(* IEC 61131-3 sources: SortJet_MasterSPS_Aufbau.fbsproj/09_Station/Stationen/Faecherwagen [301-305]/Basic_Faecherwagenstation_FB_V01_00_00.fb.st^, 19 files *)

(* ---- A_Changelog.act.st ---- *)
(* METADATA
{
	"v3Meta": {
		"objectGuid": "929bf022-d5bd-484d-b38d-56fc386ae04b"
	}
}
*)
{attribute 'excludefrombuild'}
ACTION A_Changelog
(* !!! VERSIONSÄNDERUNGEN WERDEN HIER DETAILLIERT DOKUMENTIERT !!!

- 2026-11-24 - V01_00_00: Tobias Brekerbohm
  - Erste Freigabe SortJet-Master
*)
END_ACTION

(* ---- A_ScheibenDeaktivierteStationMelden.act.st ---- *)
(* METADATA
{
	"v3Meta": {
		"objectGuid": "9787c6c4-89ac-4e67-aebe-436ca2600e9a"
	}
}
*)
ACTION A_ScheibenDeaktivierteStationMelden
// @TEXT_IMPLEMENTATION := 'ST'
//-------------------------------------------------------------------------------------------------
// DEAKTIVIERTE STATION: SCHEIBEN AN MMI MELDEN
//-------------------------------------------------------------------------------------------------
(* Hinweis:
   - Ersetzt die gleichnamige Aktion von Basic_Station_FB (auch beim Aufruf aus deren Rumpf)
   - Faecherwagenstationen melden dem MMI keine Scheiben auf der Station
*)
;
END_ACTION

(* ---- A_Schnittstelle.act.st ---- *)
(* METADATA
{
	"v3Meta": {
		"objectGuid": "4b006156-55f0-4052-a03b-8c052b439175"
	}
}
*)
ACTION A_Schnittstelle
//-------------------------------------------------------------------------------------------------
// SCHNITTSTELLE
//-------------------------------------------------------------------------------------------------

// Allgemeiner Teil: Auftrag aktiv, Stationsnummern, Fehler, Freigabe, Handfunktionen
SUPER^.A_Schnittstelle();

(* Hinweis:
   - Schnittstelle zwischen den Stationen [Transportkopplung]
*)
BasisStationsParameter.OutGlasTransport[cWAND_1].bEinlaufsensor         REF= bgFALSE;
BasisStationsParameter.OutGlasTransport[cWAND_1].bAuslaufsensor         REF= bgFALSE;
BasisStationsParameter.OutGlasTransport[cWAND_1].bBereitZumAustransport REF= bpOutBereitZumAustransport;
BasisStationsParameter.OutGlasTransport[cWAND_1].bBereitZumEintransport REF= bpOutBereitZumEintransport;
BasisStationsParameter.OutGlasTransport[cWAND_1].rGeschwindigkeit       REF= rgNULL;
END_ACTION

(* ---- A_Visu.act.st ---- *)
(* METADATA
{
	"v3Meta": {
		"objectGuid": "97dd6b9c-083d-47d5-ad19-d2fe11b9c8f1"
	}
}
*)
ACTION A_Visu
//-------------------------------------------------------------------------------------------------
// STATUS FUER DIE VISU
//-------------------------------------------------------------------------------------------------
// Allgemeiner Teil fuer alle Varianten; die Variante ergaenzt Faecherwagen, Lichtschranke und
// ihre Endlagen (abEndlage, Index = Bit der zugehoerigen Handfunktion)
IF PruefungWertImIntervall( BasisStationsParameter.stMKs.stStationsNummern.NummerSPS,
                            cERSTE_FAECHERWAGENSTATIONS_NR,
                            cLETZTE_FAECHERWAGENSTATIONS_NR )
THEN
  astgFaecherwagenstatusVisu[BasisStationsParameter.stMKs.stStationsNummern.NummerSPS].bBoxInHomePosition             := bpBoxInHomePosition;
  astgFaecherwagenstatusVisu[BasisStationsParameter.stMKs.stStationsNummern.NummerSPS].bStatusStationInBeladePosition := bpStatusStationInBeladePosition;
  astgFaecherwagenstatusVisu[BasisStationsParameter.stMKs.stStationsNummern.NummerSPS].bAuftragAktiv                  := bpAuftragAktiv;
  astgFaecherwagenstatusVisu[BasisStationsParameter.stMKs.stStationsNummern.NummerSPS].bFehler                        := BasisStationsParameter.bFehler;
  astgFaecherwagenstatusVisu[BasisStationsParameter.stMKs.stStationsNummern.NummerSPS].eStatus                        := eLetzterStatus;
  astgFaecherwagenstatusVisu[BasisStationsParameter.stMKs.stStationsNummern.NummerSPS].bRolltorOben                   := in_bRolltorGeoeffnet;
  astgFaecherwagenstatusVisu[BasisStationsParameter.stMKs.stStationsNummern.NummerSPS].bRolltorUnten                  := bpRolltorUnten;
  astgFaecherwagenstatusVisu[BasisStationsParameter.stMKs.stStationsNummern.NummerSPS].wRFID_Nummer                   := wlRFID_Nummer;
  astgFaecherwagenstatusVisu[BasisStationsParameter.stMKs.stStationsNummern.NummerSPS].abEndlage[5]                   := in_bRolltorGeoeffnet;
  astgFaecherwagenstatusVisu[BasisStationsParameter.stMKs.stStationsNummern.NummerSPS].abEndlage[6]                   := bpRolltorUnten;
END_IF
END_ACTION

(* ---- bAuftragAktiv.prop.st ---- *)
(* METADATA
{
	"v3Meta": {
		"objectGuid": "3a197e04-0bcd-4579-a4af-806c82b87acf",
		"subObjects": {
			"get": {
				"objectGuid": "bd81e771-6b2a-41b3-b424-5effe3645496"
			}
		}
	}
}
*)
PROPERTY_Get bAuftragAktiv : BOOL
VAR
END_VAR
bAuftragAktiv := bpAuftragAktiv;END_PROPERTY

(* ---- bBoxInHomePosition.prop.st ---- *)
(* METADATA
{
	"v3Meta": {
		"objectGuid": "9ae1053e-7eaa-4017-919c-7a919c9e2ca3",
		"subObjects": {
			"get": {
				"objectGuid": "c7a204ff-f1d2-4f02-aa57-0c1f7686d3d7"
			}
		}
	}
}
*)
PROPERTY_Get bBoxInHomePosition : BOOL
VAR
END_VAR
bBoxInHomePosition := bpBoxInHomePosition;END_PROPERTY

(* ---- bDone.prop.st ---- *)
(* METADATA
{
	"v3Meta": {
		"objectGuid": "7e3afc40-fd10-411a-82e2-c2f76dbe13b7",
		"subObjects": {
			"get": {
				"objectGuid": "a4174cb2-9640-462a-838e-1c212c18065f"
			}
		}
	}
}
*)
PROPERTY_Get bDone : BOOL
VAR
END_VAR
bDone := bpDone;END_PROPERTY

(* ---- bErzwingeAusschleusen.prop.st ---- *)
(* METADATA
{
	"v3Meta": {
		"objectGuid": "4cee021b-c5d5-4f3b-aa29-0070cbf1b16c",
		"subObjects": {
			"get": {
				"objectGuid": "1eace140-85af-4621-b197-e1bb9b84e0ab"
			}
		}
	}
}
*)
PROPERTY_Get bErzwingeAusschleusen : BOOL
VAR
END_VAR
bErzwingeAusschleusen := bpErzwingeAusschleusen;END_PROPERTY

(* ---- bErzwingeEinschleusen.prop.st ---- *)
(* METADATA
{
	"v3Meta": {
		"objectGuid": "82a9f007-64ac-4edb-aa26-a15d51300ac1",
		"subObjects": {
			"get": {
				"objectGuid": "2fa276e3-c875-4651-a2ef-8e71ffca1126"
			}
		}
	}
}
*)
PROPERTY_Get bErzwingeEinschleusen : BOOL
VAR
END_VAR
bErzwingeEinschleusen := bpErzwingeEinschleusen;END_PROPERTY

(* ---- bFehler.prop.st ---- *)
(* METADATA
{
	"v3Meta": {
		"objectGuid": "15bf96d6-b3ab-4293-98f3-daa693f44265",
		"subObjects": {
			"get": {
				"objectGuid": "7173d561-01b0-4b6a-be06-4d55a19c8095"
			}
		}
	}
}
*)
PROPERTY_Get bFehler : BOOL
VAR
END_VAR
bFehler := bpFehler;END_PROPERTY

(* ---- bMerkerEinschleusenQuittiert.prop.st ---- *)
(* METADATA
{
	"v3Meta": {
		"objectGuid": "bcf8d110-caa9-4eeb-bc74-c675be36606a",
		"subObjects": {
			"get": {
				"objectGuid": "c1b86ccc-2e67-4907-bc19-e7facae66067"
			}
		}
	}
}
*)
PROPERTY_Get bMerkerEinschleusenQuittiert : BOOL
VAR
END_VAR
bMerkerEinschleusenQuittiert := blMerkerEinschleusenQuittiert;END_PROPERTY

(* ---- bOutBereitZumAustransport.prop.st ---- *)
(* METADATA
{
	"v3Meta": {
		"objectGuid": "40e5f93b-ff00-4f78-b9f3-71c706ff1514",
		"subObjects": {
			"get": {
				"objectGuid": "2b4ba9cb-deb4-4b61-92f3-2bedee948b9f"
			}
		}
	}
}
*)
PROPERTY_Get bOutBereitZumAustransport : BOOL
VAR
END_VAR
bOutBereitZumAustransport := bpOutBereitZumAustransport;END_PROPERTY

(* ---- bOutBereitZumEintransport.prop.st ---- *)
(* METADATA
{
	"v3Meta": {
		"objectGuid": "529f8d13-9d58-45ad-9073-e242e51616b7",
		"subObjects": {
			"get": {
				"objectGuid": "d3cc3f71-1aa2-4715-8d89-65c33f83bf96"
			}
		}
	}
}
*)
PROPERTY_Get bOutBereitZumEintransport : BOOL
VAR
END_VAR
bOutBereitZumEintransport := bpOutBereitZumEintransport;END_PROPERTY

(* ---- bStarteSicherheitskreisReset.prop.st ---- *)
(* METADATA
{
	"v3Meta": {
		"objectGuid": "7955c67a-d244-4584-99f3-3105176a9532",
		"subObjects": {
			"set": {
				"objectGuid": "5bee3828-f9f0-4ff6-8bbd-7776959bfe22"
			},
			"get": {
				"objectGuid": "9fb27e5c-8dc6-4d5b-a84c-0ab66af3ee0d"
			}
		}
	}
}
*)
PROPERTY_Set bStarteSicherheitskreisReset : BOOL
VAR
END_VAR
// Anforderung vom MMI: Sicherheitsrelais der Station quittieren (nur Varianten mit eigenem Sicherheitsrelais werten aus)
IF ( bStarteSicherheitskreisReset ) THEN
  blStarteSicherheitskreisReset := TRUE;
END_IF
END_PROPERTY
PROPERTY_Get bStarteSicherheitskreisReset : BOOL
VAR
END_VAR
bStarteSicherheitskreisReset := blStarteSicherheitskreisReset;END_PROPERTY

(* ---- bStatusStationInBeladePosition.prop.st ---- *)
(* METADATA
{
	"v3Meta": {
		"objectGuid": "eab3fc30-cc6a-4cd0-aec6-31304c5c3cf5",
		"subObjects": {
			"get": {
				"objectGuid": "60b50eeb-6437-4f6f-8457-25ffb0000fb6"
			}
		}
	}
}
*)
PROPERTY_Get bStatusStationInBeladePosition : BOOL
VAR
END_VAR
bStatusStationInBeladePosition := bpStatusStationInBeladePosition;END_PROPERTY

(* ---- eStatus.prop.st ---- *)
(* METADATA
{
	"v3Meta": {
		"objectGuid": "92db7dc4-312f-4428-bfc2-64074944f030",
		"subObjects": {
			"get": {
				"objectGuid": "7ce800a1-a9b6-46cc-8fc0-210810cb33c8"
			}
		}
	}
}
*)
PROPERTY_Get eStatus : eLetzter_FW_Status
VAR
END_VAR
eStatus := eLetzterStatus;END_PROPERTY

(* ---- Rolltor.act.st ---- *)
(* METADATA
{
	"v3Meta": {
		"objectGuid": "7f06bdd7-dd30-4f23-890c-64b08d194069"
	}
}
*)
ACTION Rolltor
// ROLLTOR (alle Varianten, Option stStationsAufbau.bRolltor)
// ROLLTOR HOCH
// ROLLTOR HOCH

IF blRolltorAuf THEN
  CASE steplRolltorAuf OF
    // ROLLER DOOR UP  ============================
    STEP_0_E:
      blRolltorAufDone := FALSE;
      tonlZeitRunterfahren(IN := FALSE);
      tonlZeitHochfahren(IN := FALSE);
      tonlUeberwachungRolltor(IN := FALSE);
      tonlRolltorOeffnenSchliesen(IN := FALSE);

      // Schließer: TRUE = Rolltor geöffnet -> nur fahren, wenn NICHT geöffnet
      IF (NOT in_bRolltorGeoeffnet) AND BasisStationsParameter.stMKs.stStationsAufbau.bRolltor THEN
        steplRolltorAuf := STEP_5_E;
      ELSE
        steplRolltorAuf := STEP_1000_E;
      END_IF

    // ROLLTOR HOCH  ============================
    STEP_5_E:
      out_bRolltorAuf := TRUE;
      out_bRolltorAb  := FALSE;
      tonlZeitHochfahren(IN := TRUE, PT := t#60s);
      steplRolltorAuf := STEP_10_E;

    // ROLLTOR HOCH  ============================
    STEP_10_E:
      // Überwachung läuft, solange das Tor noch NICHT geöffnet ist
      tonlUeberwachungRolltor( IN := NOT in_bRolltorGeoeffnet, PT := cZEIT_UEBERWACHUNG_ROLLTOR );
      // Endlage "geöffnet" entprellen
      tonlRolltorOeffnenSchliesen( IN := in_bRolltorGeoeffnet, PT := T#500MS );
      tonlZeitHochfahren(IN := TRUE, PT := t#60s);

      IF tonlRolltorOeffnenSchliesen.Q THEN
        out_bRolltorAuf := FALSE;
        wlZeitHochfahren := TIME_TO_WORD(tonlZeitHochfahren.ET);
        tlZeitHochfahren := tonlZeitHochfahren.ET;
        tonlZeitHochfahren(IN := FALSE);
        steplRolltorAuf := STEP_1000_E;
      END_IF

      // Fehler:
      //   - Zeitliche Überwachung Rolltor
      IF tonlUeberwachungRolltor.Q THEN
        out_bRolltorAuf := FALSE;
        wpFehlerNr := cMELDUNG_FAECHERWAGEN_UEBERWACHUNG_ROLLTOR_OEFFNEN;
        SpsError( eFehler_Station,
                  wpFehlerNr,
                  BasisStationsParameter.stMKs.stStationsNummern.NummerIntern,
                  AutomatikkreisBestimmen(BasisStationsParameter.stMKs.stStationsNummern.NummerSPS),
                  BasisStationsParameter.awFehlerInformationen );

        steplRolltorAuf := STEP_900_E;
      END_IF

    // ROLLTOR HOCH  ============================
    STEP_900_E:
      out_bRolltorAb  := FALSE;
      out_bRolltorAuf := FALSE;
      BasisStationsParameter.bFehler := TRUE;

    // ROLLTOR HOCH  ============================
    STEP_1000_E:
      blRolltorAufDone := TRUE;

  // ROLLTOR HOCH  ============================
  END_CASE
ELSE

  IF ( steplRolltorAuf > STEP_0_E ) THEN
    out_bRolltorAuf  := FALSE;
    steplRolltorAuf  := STEP_0_E;
    blRolltorAufDone := FALSE;
    tonlZeitRunterfahren(IN := FALSE);
    tonlZeitHochfahren(IN := FALSE);
    tonlUeberwachungRolltor( IN := FALSE );
    tonlRolltorOeffnenSchliesen( IN := FALSE );
  END_IF

END_IF

// *********************************************************************************
// ROLLTOR RUNTER
// *********************************************************************************
IF blRolltorAb AND blRolltorAbFreigabe // Variante gibt das Schliessen frei (z.B. Lineareinheit aus dem Bereich des Rolltors)
THEN
  CASE steplRolltorAb OF
    // ROLLTOR RUNTER ============================
    STEP_0_E:
      blRolltorAbDone := FALSE;
      tonlZeitRunterfahren(IN := FALSE);
      tonlZeitHochfahren(IN := FALSE);
      tonlUeberwachungRolltor( IN := FALSE );
      tonlRolltorOeffnenSchliesen( IN := FALSE );

      IF( bpRolltorUnten OR  (NOT BasisStationsParameter.stMKs.stStationsAufbau.bRolltor))THEN
        steplRolltorAb := STEP_1000_E;
      ELSE
        steplRolltorAb := STEP_5_E;
      END_IF

    // ROLLTOR RUNTER ============================
    STEP_5_E:
      out_bRolltorAb  := TRUE;
      out_bRolltorAuf := FALSE;
      tonlZeitRunterfahren(IN := TRUE, PT := t#60s);
      tonlZeitHochfahren(IN := FALSE);
      tonlUeberwachungRolltor( IN := FALSE );
      tonlRolltorOeffnenSchliesen( IN := FALSE );
      steplRolltorAb := STEP_10_E;

    // ROLLTOR RUNTER ============================
    STEP_10_E:
      tonlUeberwachungRolltor( IN := NOT bpRolltorUnten, PT := cZEIT_UEBERWACHUNG_ROLLTOR );
      tonlRolltorOeffnenSchliesen( IN := bpRolltorUnten, PT := t#600ms );
      tonlZeitRunterfahren(IN := TRUE, PT := t#60s);

      IF tonlRolltorOeffnenSchliesen.Q THEN
        out_bRolltorAb  := FALSE;
        wlZeitRunterfahren := TIME_TO_WORD(tonlZeitRunterfahren.ET);
        tlZeitRunterfahren := tonlZeitRunterfahren.ET;
        tonlZeitRunterfahren(IN := FALSE);
        steplRolltorAb := STEP_1000_E;
      END_IF

      // Fehler:
      //   - Zeitliche Überwachung Rolltor, Abrollsicherung (Variante)
      IF tonlUeberwachungRolltor.Q OR blRolltorAbBlockiert THEN
        out_bRolltorAb := FALSE;
        wpFehlerNr := cMELDUNG_FAECHERWAGEN_UEBERWACHUNG_ROLLTOR_SCHLIESSEN;
        SpsError( eFehler_Station,
                  wpFehlerNr,
                  BasisStationsParameter.stMKs.stStationsNummern.NummerIntern,
                  AutomatikkreisBestimmen(BasisStationsParameter.stMKs.stStationsNummern.NummerSPS),
                  BasisStationsParameter.awFehlerInformationen );

        steplRolltorAb := STEP_900_E;
      END_IF

    // ROLLTOR RUNTER ============================
    STEP_900_E:
      out_bRolltorAb  := FALSE;
      out_bRolltorAuf := FALSE;
      BasisStationsParameter.bFehler := TRUE;

    // ROLLTOR RUNTER ============================
    STEP_1000_E:
      blRolltorAbDone := TRUE;

  // ROLLTOR RUNTER ============================
  END_CASE
ELSE

  IF steplRolltorAb > STEP_0_E THEN
    out_bRolltorAb  := FALSE;
    steplRolltorAb  := STEP_0_E;
    blRolltorAbDone := FALSE;
    tonlZeitRunterfahren(IN := FALSE);
    tonlZeitHochfahren(IN := FALSE);
    tonlUeberwachungRolltor( IN := FALSE );
    tonlRolltorOeffnenSchliesen( IN := FALSE );
  END_IF

END_IF
END_ACTION

(* ---- wFehlerNr.prop.st ---- *)
(* METADATA
{
	"v3Meta": {
		"objectGuid": "d72a7e2c-ee9d-4212-8954-25c76c264f34",
		"subObjects": {
			"get": {
				"objectGuid": "7e752f24-260c-4625-8435-b2c10551a2a8"
			}
		}
	}
}
*)
PROPERTY_Get wFehlerNr : WORD
VAR
END_VAR
wFehlerNr := wpFehlerNr;END_PROPERTY

(* ---- wRFID_Nummer_Schreiben.prop.st ---- *)
(* METADATA
{
	"v3Meta": {
		"objectGuid": "61bac579-e653-41b2-b8f0-3212942feb17",
		"subObjects": {
			"set": {
				"objectGuid": "2c0cfeca-c808-44fa-9f3f-5faac4060747"
			},
			"get": {
				"objectGuid": "9b84b645-b409-4691-950a-aea1dfb88055"
			}
		}
	}
}
*)
PROPERTY_Set wRFID_Nummer_Schreiben : WORD
VAR
END_VAR
// Neue Nummer fuer den RFID-Chip; die Variante schreibt bei steigender Flanke (Wert > 0)
wlRFID_Nummer_Schreiben := wRFID_Nummer_Schreiben;
END_PROPERTY
PROPERTY_Get wRFID_Nummer_Schreiben : WORD
VAR
END_VAR
wRFID_Nummer_Schreiben := wlRFID_Nummer_Schreiben;END_PROPERTY
